KUKA KRL program: Main.src

&ACCESS RVP
&REL 1
&PARAM TEMPLATE = C:\KRC\Roboter\Template\vorgabe
&PARAM EDITMASK = *
DEF Main ( )

; External program calls:
EXT WeldPair1()
EXT WeldPair2()
EXT WeldPair3()
EXT DoWeld()

EXT BAS (BAS_COMMAND :IN,REAL :IN )


; GLOBAL INTERRUPT DECL 3 WHEN $STOPMESS==TRUE DO IR_STOPM ( )
; INTERRUPT ON 3

;FOLD Initialise and set default speed
BAS (#INITMOV,0)
BAS (#VEL_PTP,100)
BAS (#ACC_PTP,20)
$VEL.CP=0.2
BAS (#TOOL,0)
BAS (#BASE,0)
;ENDFOLD

;;FOLD STARTPOS
;$BWDSTART = FALSE
;PDAT_ACT = PDEFAULT
;BAS(#PTP_DAT)
;FDAT_ACT = {TOOL_NO 0,BASE_NO 0,IPO_FRAME #BASE}
;BAS(#FRAMES)
;;ENDFOLD

$ADVANCE = 5

;FOLD ---- Quickly skip BCO ----
; PTP $AXIS_ACT
;ENDFOLD

;FOLD ---- GO HOME ----
; PTP {A1 0.000, A2 -90.000, A3 90.000, A4 0.000, A5 0.000, A6 0.000, E1 0, E2 0, E3 0, E4 0, E5 0, E6 0}
;ENDFOLD


; Program generated by VerticalBot Studio for KUKA KR 120 R2900 extra on 25/10/2026 12:00:00
; Using nominal kinematics.
; ---- Setting reference (Base) ----
$BASE = {FRAME: X 1482.740,Y 183.671,Z -402.167,A 6.534,B 0.000,C 0.000}
; --------------------------
; ---- Setting tool (TCP) ----
$TOOL = {FRAME: X 0.270,Y 0.000,Z 1049.990,A 0.000,B -90.000,C 0.000}
; --------------------------
PTP {A1 -0.00000,A2 -81.64360,A3 70.78240,A4 0.00000,A5 92.14690,A6 0.00000}
WeldPair1()
WeldPair2()
WeldPair3()
PTP {A1 -0.00000,A2 -81.64360,A3 70.78240,A4 0.00000,A5 92.14690,A6 0.00000}
END
